Fanuc KAREL source: KT00541.KL

PROGRAM KT00541
%NOLOCKGROUP
VAR
  P1: JOINTPOS
  P2: XYZWPR
  OUT: XYZWPREXT
BEGIN
    P2.Y = 2.0
  OUT = P1 : P2
END KT00541
